FUNCTION_BLOCK ResetSequence (* CAT Function Block Type *)
  (* Standard: 61499-2 *)
  (* Version 0.0, 10/23/2026, Schneider Electric, template *)
  PACKAGE Main;
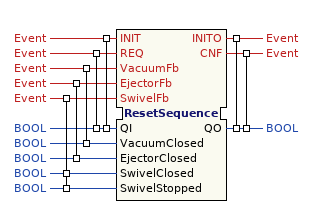
  EVENT_INPUT
    INIT WITH QI; (* Initialization Request *)
    REQ WITH QI; (* Normal Execution Request *)
    VacuumFb WITH VacuumClosed;
    EjectorFb WITH EjectorClosed;
    SwivelFb WITH SwivelClosed, SwivelStopped;
  END_EVENT
  EVENT_OUTPUT
    INITO WITH QO; (* Initialization Confirm *)
    CNF WITH QO; (* Execution Confirmation *)
  END_EVENT
  VAR_INPUT
    QI : BOOL; (* Input event qualifier *)
    VacuumClosed : BOOL;
    EjectorClosed : BOOL;
    SwivelClosed : BOOL;
    SwivelStopped : BOOL;
  END_VAR
  VAR_OUTPUT
    QO : BOOL; (* Output event qualifier *)
  END_VAR
  FBS
    ResetSeq : SeqHead(PermStart := TRUE);
    RS1_TakeOver : SeqStep(TransStepId := 2);
    RS_End : SeqTerminate;
    Consts : ANY2ANY_25FC8D56FEEDC9B5(IN1 := TRUE, IN2 := 1, IN3 := 2, IN4 := 0); {SET_ATTRIBUTE(Configuration.GenericFBType.InterfaceParams, Runtime.Standard#CNT:=4;IN${CNT$}:BOOL,INT,INT,INT;OUT${CNT$}:VTQBOOL,VTQINT,VTQINT,VTQINT)}
    RS3_EjectorBack : SeqStep(TransStepId := 4);
    RS2_VacuumOff : SeqStep(TransStepId := 3);
    RS4_SwivelHome : SeqStep(TransStepId := 5);
    RS5_SwivelOffMag : SeqStep(TransStepId := 6);
    RS6_SwivelParkStop : SeqStep(TransStepId := 7);
    OwnerFb : SYMLINKMULTIVARDST_105A0442B8CC61A96(NAME1 := 'RES0.Distribution.Vacuum.sc.progLocal', NAME2 := 'RES0.Distribution.Ejector.sc.progLocal', NAME3 := 'RES0.Distribution.Swivel.sc.progLocal', QI := TRUE); {SET_ATTRIBUTE(Configuration.GenericFBType.InterfaceParams, Runtime.System#I:=3;VALUE${I$}:VTQBOOL,VTQBOOL,VTQBOOL)}
    TakeOverCmd : SYMLINKMULTIVARSRC_105A0442B8CC61A96(QI := TRUE, NAME1 := 'RES0.Distribution.Vacuum.sc.progLocalSel', NAME2 := 'RES0.Distribution.Ejector.sc.progLocalSel', NAME3 := 'RES0.Distribution.Swivel.sc.progLocalSel'); {SET_ATTRIBUTE(Configuration.GenericFBType.InterfaceParams, Runtime.System#I:=3;VALUE${I$}:VTQBOOL,VTQBOOL,VTQBOOL)}
    EjectorBackCmd : SYMLINKMULTIVARSRC_18556BCA74EA878F1(QI := TRUE, NAME1 := 'RES0.Distribution.Ejector.sc.lsp'); {SET_ATTRIBUTE(Configuration.GenericFBType.InterfaceParams, Runtime.System#I:=1;VALUE${I$}:VTQINT)}
    VacuumOffCmd : SYMLINKMULTIVARSRC_18556BCA74EA878F1(QI := TRUE, NAME1 := 'RES0.Distribution.Vacuum.sc.lsp'); {SET_ATTRIBUTE(Configuration.GenericFBType.InterfaceParams, Runtime.System#I:=1;VALUE${I$}:VTQINT)}
    SwivelHomeCmd : SYMLINKMULTIVARSRC_18556BCA74EA878F1(QI := TRUE, NAME1 := 'RES0.Distribution.Swivel.sc.lsp'); {SET_ATTRIBUTE(Configuration.GenericFBType.InterfaceParams, Runtime.System#I:=1;VALUE${I$}:VTQINT)}
    AllLocal : AND_550FE6D62F509EB3(IN3 := TRUE); {SET_ATTRIBUTE(Configuration.GenericFBType.InterfaceParams, Runtime.Standard#CNT:=3;OUT:BOOL)}
    ArmOffMag : NOT_42C76073DCEB1A7A; {SET_ATTRIBUTE(Configuration.GenericFBType.InterfaceParams, Runtime.Standard#CNT:=1;OUT${CNT$}:BOOL)}
    SwivelOutCmd : SYMLINKMULTIVARSRC_18556BCA74EA878F1(QI := TRUE, NAME1 := 'RES0.Distribution.Swivel.sc.lsp'); {SET_ATTRIBUTE(Configuration.GenericFBType.InterfaceParams, Runtime.System#I:=1;VALUE${I$}:VTQINT)}
    SwivelStopCmd : SYMLINKMULTIVARSRC_18556BCA74EA878F1(QI := TRUE, NAME1 := 'RES0.Distribution.Swivel.sc.lsp'); {SET_ATTRIBUTE(Configuration.GenericFBType.InterfaceParams, Runtime.System#I:=1;VALUE${I$}:VTQINT)}
  END_FBS
  EVENT_CONNECTIONS
    INIT TO Consts.REQ;
    Consts.CNF TO ResetSeq.REQ_PERM;
    Consts.CNF TO TakeOverCmd.INIT;
    Consts.CNF TO VacuumOffCmd.INIT;
    Consts.CNF TO EjectorBackCmd.INIT;
    Consts.CNF TO SwivelHomeCmd.INIT;
    Consts.CNF TO SwivelOutCmd.INIT;
    Consts.CNF TO SwivelStopCmd.INIT;
    Consts.CNF TO OwnerFb.INIT;
    OwnerFb.CNF TO AllLocal.REQ;
    AllLocal.CNF TO RS1_TakeOver.TRANS_REQ;
    RS1_TakeOver.STEP_ENTER TO TakeOverCmd.REQ;
    TakeOverCmd.CNF TO AllLocal.REQ;
    RS2_VacuumOff.STEP_ENTER TO VacuumOffCmd.REQ;
    RS3_EjectorBack.STEP_ENTER TO EjectorBackCmd.REQ;
    RS4_SwivelHome.STEP_ENTER TO SwivelHomeCmd.REQ;
    EjectorBackCmd.CNF TO RS3_EjectorBack.TRANS_REQ;
    VacuumOffCmd.CNF TO RS2_VacuumOff.TRANS_REQ;
    SwivelHomeCmd.CNF TO RS4_SwivelHome.TRANS_REQ;
    VacuumFb TO RS2_VacuumOff.TRANS_REQ;
    EjectorFb TO RS3_EjectorBack.TRANS_REQ;
    SwivelFb TO RS4_SwivelHome.TRANS_REQ;
    RS5_SwivelOffMag.STEP_ENTER TO SwivelOutCmd.REQ;
    SwivelOutCmd.CNF TO ArmOffMag.REQ;
    SwivelFb TO ArmOffMag.REQ;
    ArmOffMag.CNF TO RS5_SwivelOffMag.TRANS_REQ;
    RS6_SwivelParkStop.STEP_ENTER TO SwivelStopCmd.REQ;
    SwivelStopCmd.CNF TO RS6_SwivelParkStop.TRANS_REQ;
    SwivelFb TO RS6_SwivelParkStop.TRANS_REQ;
  END_CONNECTIONS
  DATA_CONNECTIONS
    Consts.OUT1 TO TakeOverCmd.VALUE1;
    Consts.OUT1 TO TakeOverCmd.VALUE2;
    Consts.OUT1 TO TakeOverCmd.VALUE3;
    Consts.OUT3 TO VacuumOffCmd.VALUE1;
    Consts.OUT3 TO EjectorBackCmd.VALUE1;
    Consts.OUT3 TO SwivelHomeCmd.VALUE1;
    Consts.OUT2 TO SwivelOutCmd.VALUE1;
    Consts.OUT4 TO SwivelStopCmd.VALUE1;
    OwnerFb.VALUE1 TO AllLocal.IN1;
    OwnerFb.VALUE2 TO AllLocal.IN2;
    AllLocal.OUT TO RS1_TakeOver.Exceeded;
    VacuumClosed TO RS2_VacuumOff.Exceeded;
    EjectorClosed TO RS3_EjectorBack.Exceeded;
    SwivelClosed TO RS4_SwivelHome.Exceeded;
    SwivelClosed TO ArmOffMag.IN1;
    ArmOffMag.OUT1 TO RS5_SwivelOffMag.Exceeded;
    SwivelStopped TO RS6_SwivelParkStop.Exceeded;
  END_CONNECTIONS
  ADAPTER_CONNECTIONS
    ResetSeq.ISeqChain TO RS1_TakeOver.ISeqChainIn;
    RS1_TakeOver.ISeqChainOut TO RS2_VacuumOff.ISeqChainIn;
    RS2_VacuumOff.ISeqChainOut TO RS3_EjectorBack.ISeqChainIn;
    RS3_EjectorBack.ISeqChainOut TO RS4_SwivelHome.ISeqChainIn;
    RS4_SwivelHome.ISeqChainOut TO RS5_SwivelOffMag.ISeqChainIn;
    RS5_SwivelOffMag.ISeqChainOut TO RS6_SwivelParkStop.ISeqChainIn;
    RS6_SwivelParkStop.ISeqChainOut TO RS_End.ISeqChainIn;
  END_CONNECTIONS
END_FUNCTION_BLOCK
